ABB RAPID module: ManyMoves.mod

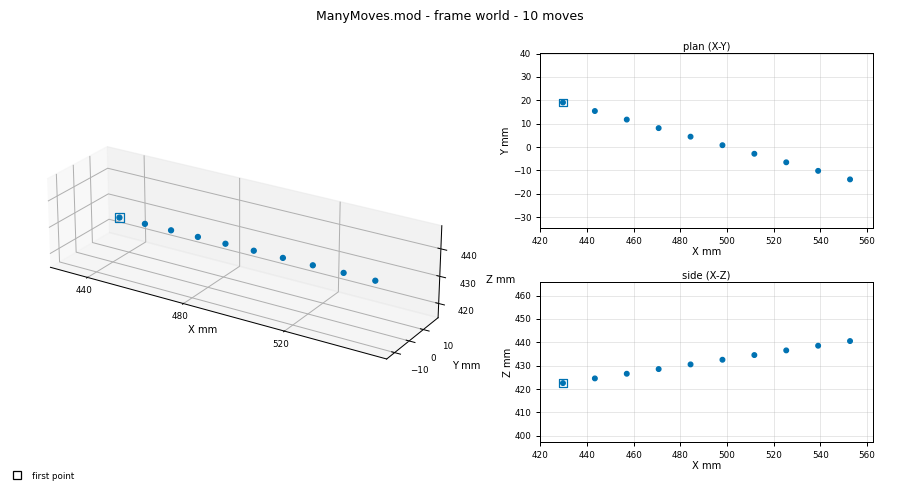
[picture p0: tool path of ManyMoves.mod in frame world, 10 of 40 moves have a stored position in this frame; points joined in program order, loops and branches not executed]
%%%
  VERSION:1
  LANGUAGE:ENGLISH
%%%
MODULE MOD_ManyMoves

    ! -------------------------------
    ! Define customized variables here
    ! ...

	! Tool variables:
	PERS tooldata ToolS := [TRUE,[[10.000,20.000,150.000],[1.00000000,0.00000000,0.00000000,0.00000000]],[1,[0,0,20],[1,0,0,0],0,0,0.005]];

	! Reference variables:
	PERS wobjdata FrameS := [FALSE, TRUE, "", [[0,0,0],[1,0,0,0]],[[1234.570,-98.765,50.500],[0.96592583,0.00000000,0.00000000,0.25881905]]];

	PROC Main()
		ConfJ \On;
		ConfL \Off;
		! Program generated by RoboDK v6.0.7 for ABB IRB 260 on XX/XX/XXXX 18:00:00
		! Using nominal kinematics.
		MoveAbsJ [[10.000000,-20.000000,50.000000,30.000000,0.000000,0.000000],[9E+09,9E+09,9E+09,9E+09,9E+09,9E+09]],v500,z1,ToolS \WObj:=FrameS;
		MoveL [[-638.084,504.480,372.034],[0.37410804,0.28584607,0.85365954,-0.22271191],[0,0,0,0],[9E+09,9E+09,9E+09,9E+09,9E+09,9E+09]],v500,z1,ToolS \WObj:=FrameS;
		MoveAbsJ [[30.000000,25.000000,80.000000,-45.000000,0.000000,0.000000],[9E+09,9E+09,9E+09,9E+09,9E+09,9E+09]],v500,z1,ToolS \WObj:=FrameS;
		MoveL CalcRobT([[10.000000,-20.000000,50.000000,30.000000,0.000000,0.000000],[9E+09,9E+09,9E+09,9E+09,9E+09,9E+09]],ToolS \WObj:=FrameS),v500,z1,ToolS \WObj:=FrameS;
		MoveAbsJ [[10.000000,-20.000000,50.000000,30.000000,0.000000,0.000000],[9E+09,9E+09,9E+09,9E+09,9E+09,9E+09]],v500,z1,ToolS \WObj:=FrameS;
		MoveL [[-628.084,494.480,374.034],[0.37410804,0.28584607,0.85365954,-0.22271191],[0,0,0,0],[9E+09,9E+09,9E+09,9E+09,9E+09,9E+09]],v500,z1,ToolS \WObj:=FrameS;
		MoveAbsJ [[30.000000,25.000000,80.000000,-45.000000,0.000000,0.000000],[9E+09,9E+09,9E+09,9E+09,9E+09,9E+09]],v500,z1,ToolS \WObj:=FrameS;
		MoveL CalcRobT([[10.000000,-20.000000,50.000000,30.000000,0.000000,0.000000],[9E+09,9E+09,9E+09,9E+09,9E+09,9E+09]],ToolS \WObj:=FrameS),v500,z1,ToolS \WObj:=FrameS;
		MoveAbsJ [[10.000000,-20.000000,50.000000,30.000000,0.000000,0.000000],[9E+09,9E+09,9E+09,9E+09,9E+09,9E+09]],v500,z1,ToolS \WObj:=FrameS;
		MoveL [[-618.084,484.480,376.034],[0.37410804,0.28584607,0.85365954,-0.22271191],[0,0,0,0],[9E+09,9E+09,9E+09,9E+09,9E+09,9E+09]],v500,z1,ToolS \WObj:=FrameS;
		MoveAbsJ [[30.000000,25.000000,80.000000,-45.000000,0.000000,0.000000],[9E+09,9E+09,9E+09,9E+09,9E+09,9E+09]],v500,z1,ToolS \WObj:=FrameS;
		MoveL CalcRobT([[10.000000,-20.000000,50.000000,30.000000,0.000000,0.000000],[9E+09,9E+09,9E+09,9E+09,9E+09,9E+09]],ToolS \WObj:=FrameS),v500,z1,ToolS \WObj:=FrameS;
		MoveAbsJ [[10.000000,-20.000000,50.000000,30.000000,0.000000,0.000000],[9E+09,9E+09,9E+09,9E+09,9E+09,9E+09]],v500,z1,ToolS \WObj:=FrameS;
		MoveL [[-608.084,474.480,378.034],[0.37410804,0.28584607,0.85365954,-0.22271191],[0,0,0,0],[9E+09,9E+09,9E+09,9E+09,9E+09,9E+09]],v500,z1,ToolS \WObj:=FrameS;
		MoveAbsJ [[30.000000,25.000000,80.000000,-45.000000,0.000000,0.000000],[9E+09,9E+09,9E+09,9E+09,9E+09,9E+09]],v500,z1,ToolS \WObj:=FrameS;
		MoveL CalcRobT([[10.000000,-20.000000,50.000000,30.000000,0.000000,0.000000],[9E+09,9E+09,9E+09,9E+09,9E+09,9E+09]],ToolS \WObj:=FrameS),v500,z1,ToolS \WObj:=FrameS;
		MoveAbsJ [[10.000000,-20.000000,50.000000,30.000000,0.000000,0.000000],[9E+09,9E+09,9E+09,9E+09,9E+09,9E+09]],v500,z1,ToolS \WObj:=FrameS;
		MoveL [[-598.084,464.480,380.034],[0.37410804,0.28584607,0.85365954,-0.22271191],[0,0,0,0],[9E+09,9E+09,9E+09,9E+09,9E+09,9E+09]],v500,z1,ToolS \WObj:=FrameS;
		MoveAbsJ [[30.000000,25.000000,80.000000,-45.000000,0.000000,0.000000],[9E+09,9E+09,9E+09,9E+09,9E+09,9E+09]],v500,z1,ToolS \WObj:=FrameS;
		MoveL CalcRobT([[10.000000,-20.000000,50.000000,30.000000,0.000000,0.000000],[9E+09,9E+09,9E+09,9E+09,9E+09,9E+09]],ToolS \WObj:=FrameS),v500,z1,ToolS \WObj:=FrameS;
		MoveAbsJ [[10.000000,-20.000000,50.000000,30.000000,0.000000,0.000000],[9E+09,9E+09,9E+09,9E+09,9E+09,9E+09]],v500,z1,ToolS \WObj:=FrameS;
		MoveL [[-588.084,454.480,382.034],[0.37410804,0.28584607,0.85365954,-0.22271191],[0,0,0,0],[9E+09,9E+09,9E+09,9E+09,9E+09,9E+09]],v500,z1,ToolS \WObj:=FrameS;
		MoveAbsJ [[30.000000,25.000000,80.000000,-45.000000,0.000000,0.000000],[9E+09,9E+09,9E+09,9E+09,9E+09,9E+09]],v500,z1,ToolS \WObj:=FrameS;
		MoveL CalcRobT([[10.000000,-20.000000,50.000000,30.000000,0.000000,0.000000],[9E+09,9E+09,9E+09,9E+09,9E+09,9E+09]],ToolS \WObj:=FrameS),v500,z1,ToolS \WObj:=FrameS;
		MoveAbsJ [[10.000000,-20.000000,50.000000,30.000000,0.000000,0.000000],[9E+09,9E+09,9E+09,9E+09,9E+09,9E+09]],v500,z1,ToolS \WObj:=FrameS;
		MoveL [[-578.084,444.480,384.034],[0.37410804,0.28584607,0.85365954,-0.22271191],[0,0,0,0],[9E+09,9E+09,9E+09,9E+09,9E+09,9E+09]],v500,z1,ToolS \WObj:=FrameS;
		MoveAbsJ [[30.000000,25.000000,80.000000,-45.000000,0.000000,0.000000],[9E+09,9E+09,9E+09,9E+09,9E+09,9E+09]],v500,z1,ToolS \WObj:=FrameS;
		MoveL CalcRobT([[10.000000,-20.000000,50.000000,30.000000,0.000000,0.000000],[9E+09,9E+09,9E+09,9E+09,9E+09,9E+09]],ToolS \WObj:=FrameS),v500,z1,ToolS \WObj:=FrameS;
		MoveAbsJ [[10.000000,-20.000000,50.000000,30.000000,0.000000,0.000000],[9E+09,9E+09,9E+09,9E+09,9E+09,9E+09]],v500,z1,ToolS \WObj:=FrameS;
		MoveL [[-568.084,434.480,386.034],[0.37410804,0.28584607,0.85365954,-0.22271191],[0,0,0,0],[9E+09,9E+09,9E+09,9E+09,9E+09,9E+09]],v500,z1,ToolS \WObj:=FrameS;
		MoveAbsJ [[30.000000,25.000000,80.000000,-45.000000,0.000000,0.000000],[9E+09,9E+09,9E+09,9E+09,9E+09,9E+09]],v500,z1,ToolS \WObj:=FrameS;
		MoveL CalcRobT([[10.000000,-20.000000,50.000000,30.000000,0.000000,0.000000],[9E+09,9E+09,9E+09,9E+09,9E+09,9E+09]],ToolS \WObj:=FrameS),v500,z1,ToolS \WObj:=FrameS;
		MoveAbsJ [[10.000000,-20.000000,50.000000,30.000000,0.000000,0.000000],[9E+09,9E+09,9E+09,9E+09,9E+09,9E+09]],v500,z1,ToolS \WObj:=FrameS;
		MoveL [[-558.084,424.480,388.034],[0.37410804,0.28584607,0.85365954,-0.22271191],[0,0,0,0],[9E+09,9E+09,9E+09,9E+09,9E+09,9E+09]],v500,z1,ToolS \WObj:=FrameS;
		MoveAbsJ [[30.000000,25.000000,80.000000,-45.000000,0.000000,0.000000],[9E+09,9E+09,9E+09,9E+09,9E+09,9E+09]],v500,z1,ToolS \WObj:=FrameS;
		MoveL CalcRobT([[10.000000,-20.000000,50.000000,30.000000,0.000000,0.000000],[9E+09,9E+09,9E+09,9E+09,9E+09,9E+09]],ToolS \WObj:=FrameS),v500,z1,ToolS \WObj:=FrameS;
		MoveAbsJ [[10.000000,-20.000000,50.000000,30.000000,0.000000,0.000000],[9E+09,9E+09,9E+09,9E+09,9E+09,9E+09]],v500,z1,ToolS \WObj:=FrameS;
		MoveL [[-548.084,414.480,390.034],[0.37410804,0.28584607,0.85365954,-0.22271191],[0,0,0,0],[9E+09,9E+09,9E+09,9E+09,9E+09,9E+09]],v500,z1,ToolS \WObj:=FrameS;
		MoveAbsJ [[30.000000,25.000000,80.000000,-45.000000,0.000000,0.000000],[9E+09,9E+09,9E+09,9E+09,9E+09,9E+09]],v500,z1,ToolS \WObj:=FrameS;
		MoveL CalcRobT([[10.000000,-20.000000,50.000000,30.000000,0.000000,0.000000],[9E+09,9E+09,9E+09,9E+09,9E+09,9E+09]],ToolS \WObj:=FrameS),v500,z1,ToolS \WObj:=FrameS;
	ENDPROC

ENDMODULE
